Fanuc KAREL source: KB00007.KL

PROGRAM KB00007
%NOLOCKGROUP
%ENVIRONMENT VECTR
VAR
  P1: POSITION
  RESULT: VECTOR
BEGIN
  RESULT = APPROACH(P1)
END KB00007
